# EPICS autosave request: soft_iocs/xds_optics/iocBoot/iocxds_optics/mono_settings.req
file monoModes_settings.req P=18ID:, MN=Mono
file pseudoMotor_settings.req P=18ID:Mono:, M=Energy
file pseudoMotor_settings.req P=18ID:Mono:, M=Offset
file pseudoMotor_settings.req P=18ID:Mono:, M=Lambda

#
